FUNCTION_BLOCK FB_Valve
VAR_INPUT
    R       : Bool;
    nSpeed  : Int;  // speed
END_VAR
VAR
    sTimer  : TON;
    sbDone  : Bool;
END_VAR

If R Then
    sTimer
        (
         IN := True,
         PT := T#5S,
         Q  => sbDone
         );
End_If

METHOD M_Reset : Bool
VAR_INPUT
    bForce  : Bool;
END_VAR
VAR
    x       : Int;
END_VAR
x           := 0;
M_Reset     := True;
END_METHOD

END_FUNCTION_BLOCK

(* stored: Version 1.1.0.1, ProductVersion 3.1.4024.12
   POU FB_Valve: Id {11111111-2222-3333-4444-555555555555}, SpecialFunc None
   Method M_Reset: Id {aaaaaaaa-2222-3333-4444-555555555555} *)
